// TIA Portal V20 export
TYPE "WT2_Vd_Status_1_UDT"
   STRUCT
      iHandshake : Int;
      Fehler : Struct
         bE0000_KonfigFehler : Bool;
         bE0001_VerbundMasterAusg : Bool;
         bE0002_NotstoppPHDFehler : Bool;
         bE0003_ExternFehler : Bool;
         bE0004_TDruckFehler : Bool;
         bE0005_PDruckFehler : Bool;
         bE0006_PSaugFehler : Bool;
         bE0007_TMotorFehler : Bool;
         bE0008_TSHMinSaugFehler : Bool;
         bE0009_TSHMinDruckFehler : Bool;
         bE0010_LuefterFehler : Bool;
         bE0011_Reserviert : Bool;
         bE0012_PhasenFehler : Bool;
         bE0013_MotorFehler : Bool;
         bE0014_LSAusloesung : Bool;
         bE0015_POeldiffStillstand : Bool;
         bE0016_POeldiffBetrieb : Bool;
         bE0017_TOelMaxFehler : Bool;
         bE0018_OElniveauOA : Bool;
         bE0019_OElniveauVd : Bool;
         bE0020_OElStroemung : Bool;
         bE0021_POelfilterBetrieb : Bool;
         bE0022_TLagerDEFehler : Bool;
         bE0023_TLager_NDEFehler : Bool;
         bE0024_Reserviert : Bool;
         bE0025_Reserviert : Bool;
         bE0026_Reserviert : Bool;
         bE0027_PSaugOverrange : Bool;
         bE0028_PPsZuTief : Bool;
         bE0029_Oelpumpe : Bool;
         bE0030_Leistungsschieber : Bool;
         bE0031_PoPsZuTief : Bool;
         bE0032_StartdruckZuHoch : Bool;
         bE0033_POelfilterStillstand : Bool;
         bE0034_PoPMinFehler : Bool;
         bE0035_Startoeldruck : Bool;
         bE0036_TDruckGradient : Bool;
         bE0037_OelflussVerdichter : Bool;
         bE0038_KeineGasfoerderung : Bool;
         bE0039_PZwDruck : Bool;
         bE0040_TZwDruck : Bool;
         bE0041_TSHMinZwDruck : Bool;
         bE0042_POeldiffMax : Bool;
         bE0043_PPsMax : Bool;
         bE0044_OelkhlungTop : Bool;
         bE0045_PPzZuTeif : Bool;
         bE0046_PPzMax : Bool;
         bE0047_PPsZuTief : Bool;
         bE0048_FluessigSchlag : Bool;
         bE0049_Reserviert : Bool;
         bE0050_Reserviert : Bool;
         bE0051_Reserviert : Bool;
         bE0052_Reserviert : Bool;
         bE0053_Reserviert : Bool;
         bE0054_Reserviert : Bool;
         bE0055_Reserviert : Bool;
         bE0056_Reserviert : Bool;
         bE0057_Reserviert : Bool;
         bE0058_Reserviert : Bool;
         bE0059_Reserviert : Bool;
         bE0060_Reserviert : Bool;
         bE0061_Reserviert : Bool;
         bE0062_Reserviert : Bool;
         bE0063_KaeltekreisMasterAusgefa : Bool;
         bE0064_Reserviert : Bool;
         bE0065_KaelteKreisInvUngueltig : Bool;
         bE0066_OelkreisMasterAusgefa : Bool;
         bE0067_Reserviert : Bool;
         bE0068_OelKreisInvUngueltig : Bool;
         bE0069_SchmierdruckMin : Bool;
         bE0070_PPoMax : Bool;
         bE0071_Haupt_OeldruckMin : Bool;
         bE0072_Reserviert : Bool;
         bE0073_Reserviert : Bool;
         bE0074_Reserviert : Bool;
         bE0075_TZylinderkopfFehler : Bool;
         bE0076_VerdampferpumpeFehlerBet : Bool;
         bE0077_VerdampferpumpeFehlerSti : Bool;
         bE0078_NivHDAbschHochFehler : Bool;
         bE0079_NivEconomiserHochFehler : Bool;
         bE0080_Reserviert : Bool;
         bE0081_KonfFehlerKkStart_Stopp : Bool;
         bE0082_HDVerdAusgefallen : Bool;
         bE0083_NDVerdAusgefallen : Bool;
         bE0084_KeinStartbefehlKonf : Bool;
         bE0085_PzPsMax : Bool;
         bE0086_Reserviert : Bool;
         bE0087_VibraSwitchAusg : Bool;
         bE0088_TOelabschMax : Bool;
         bE0089_TOelMin : Bool;
         bE0090_Reserviert : Bool;
         bE0091_NDAbschNivHoch : Bool;
         bE0092_Sekundaerschieber : Bool;
         bE0093_Reserviert : Bool;
         bE0094_KonfigFehlerAbsKuehls : Bool;
         bE0095_Reserviert : Bool;
         bE0096_OelnivKGHhoch : Bool;
         bE0097_KonfigFehlerDIPrio : Bool;
         bE0098_Reserviert : Bool;
         bE0099_Reserviert : Bool;
         bE0100_Reserviert : Bool;
         bE0101_KonfigFehlerDrehzahl : Bool;
         bE0102_Reserviert : Bool;
         bE0103_PSaugHoch : Bool;
         bE0104_KonfigFehlerMotorleist : Bool;
         bE0105_FehlerEinsatzdiagr : Bool;
         bE0106_Reserviert : Bool;
         bE0107_Reserviert : Bool;
         bE0108_Reserviert : Bool;
         bE0109_MotorfehlerNotAusTest : Bool;
         bE0110_StirnspHauptrotorZGross : Bool;
         bE0111_StirnspHautprotorZKlein : Bool;
         bE0112_StirnspNebenrotorZGross : Bool;
         bE0113_StirnspNebenrotorZKlein : Bool;
         bE0114_THauptrotorDS : Bool;
         bE0115_THauptrotorSS : Bool;
         bE0116_TNebenrotorDS : Bool;
         bE0117_TNebenrotorSS : Bool;
         bE0118_FlSchlagFehlerSensor : Bool;
         bE0119_OelstoppventilFehler : Bool;
         bE0120_Reserviert : Bool;
         bE0121_Reserviert : Bool;
         bE0122_Reserviert : Bool;
         bE0123_Reserviert : Bool;
         bE0124_Reserviert : Bool;
         bE0125_Reserviert : Bool;
         bE0126_Reserviert : Bool;
         bE0127_Reserviert : Bool;
      END_STRUCT;
      Alarm : Struct
         bA1000_Reserviert : Bool;
         bA1001_VerbundMasterAusg : Bool;
         bA1002_Reserviert : Bool;
         bA1003_Reserviert : Bool;
         bA1004_TDruck : Bool;
         bA1005_PDruck : Bool;
         bA1006_Reserviert : Bool;
         bA1007_TMotor : Bool;
         bA1008_TSHMinSaug : Bool;
         bA1009_TSHMinDruck : Bool;
         bA1010_Reserviert : Bool;
         bA1011_Reserviert : Bool;
         bA1012_Reserviert : Bool;
         bA1013_Reserviert : Bool;
         bA1014_Reserviert : Bool;
         bA1015_Reserviert : Bool;
         bA1016_POeldiff_Betrieb : Bool;
         bA1017_TOelmax : Bool;
         bA1018_OelniveauOA : Bool;
         bA1019_Reserviert : Bool;
         bA1020_Reserviert : Bool;
         bA1021_POelfilterBetrieb : Bool;
         bA1022_TLagerDE : Bool;
         bA1023_TLagerNDE : Bool;
         bA1024_OelniveauOA_hoch : Bool;
         bA1025_Reserviert : Bool;
         bA1026_Reserviert : Bool;
         bA1027_PSaugOverrange : Bool;
         bA1028_PPszutief : Bool;
         bA1029_Reserviert : Bool;
         bA1030_Reserviert : Bool;
         bA1031_Reserviert : Bool;
         bA1032_Reserviert : Bool;
         bA1033_Reserviert : Bool;
         bA1034_PoPMin : Bool;
         bA1035_Reserviert : Bool;
         bA1036_Reserviert : Bool;
         bA1037_Reserviert : Bool;
         bA1038_Reserviert : Bool;
         bA1039_PZwDruck : Bool;
         bA1040_TZwDruck : Bool;
         bA1041_TSHminZwDruck : Bool;
         bA1042_Reserviert : Bool;
         bA1043_PPsmax : Bool;
         bA1044_Reserviert : Bool;
         bA1045_PPzzutief : Bool;
         bA1046_PPzmax : Bool;
         bA1047_PPszutief2 : Bool;
         bA1048_FluessigSchlag : Bool;
         bA1049_NDPendel : Bool;
         bA1050_TOelMin : Bool;
         bA1051_Reserviert : Bool;
         bA1052_OelheizungOA : Bool;
         bA1053_TSaug : Bool;
         bA1054_PSauglimit : Bool;
         bA1055_PDrucklimit : Bool;
         bA1056_LastabwurfMotorstrom : Bool;
         bA1057_MinLeistungnErr : Bool;
         bA1058_MaxLeistungnErr : Bool;
         bA1059_BalanceFNorm : Bool;
         bA1060_PrimaerschMaxNErr : Bool;
         bA1061_LastabwurfMotorleistung : Bool;
         bA1062_OelheizungKGH : Bool;
         bA1063_KaeltekreisMasterAusgef : Bool;
         bA1064_KaeltekreisSlaveAusgef : Bool;
         bA1065_Reserviert : Bool;
         bA1066_Reserviert : Bool;
         bA1067_OelkreisSlaveAusgef : Bool;
         bA1068_Reserviert : Bool;
         bA1069_SchmierdruckMin : Bool;
         bA1070_PPoMax : Bool;
         bA1071_HauptOeldruckMin : Bool;
         bA1072_Oelnachspeisung : Bool;
         bA1073_KdMasterAusgef : Bool;
         bA1074_VrMasterAusgef : Bool;
         bA1075_TZylinderkopf : Bool;
         bA1076_Reserviert : Bool;
         bA1077_Reserviert : Bool;
         bA1078_Reserviert : Bool;
         bA1079_Reserviert : Bool;
         bA1080_KdMasterAusef : Bool;
         bA1081_Reserviert : Bool;
         bA1082_Reserviert : Bool;
         bA1083_Reserviert : Bool;
         bA1084_Reserviert : Bool;
         bA1085_PzPsAlarm : Bool;
         bA1086_HauptMasterAusgef : Bool;
         bA1087_Reserviert : Bool;
         bA1088_TOelabschMaxAlarm : Bool;
         bA1089_TOelMinAlarm : Bool;
         bA1090_OelpumpePendelalarm : Bool;
         bA1091_Reserviert : Bool;
         bA1092_Reserviert : Bool;
         bA1093_TOelMinAlarmKGH : Bool;
         bA1094_Reserviert : Bool;
         bA1095_TZwDruckSaugHDAlarm : Bool;
         bA1096_OelniveauKGHHoch : Bool;
         bA1097_Reserviert : Bool;
         bA1098_MKaeltekrMasterAktiv : Bool;
         bA1099_MOelkreisMasterAktiv : Bool;
         "bA1100_Objekt-ID mehrfach vorhanden" : Bool;
         bA1101_Reserviert : Bool;
         bA1102_RekalibrierungMinNDurchg : Bool;
         bA1103_Reserviert : Bool;
         bA1104_Reserviert : Bool;
         bA1105_AlarmEinsatzdiagr : Bool;
         bA1106_AlarmEcoNivEndsch : Bool;
         bA1107_OelnachspDVrGesp : Bool;
         bA1108_OerektDVrGesp : Bool;
         bA1109_NotAusTestFehlgeschl : Bool;
         bA1110_StirnspHauptrotorZGross : Bool;
         bA1111_StirnspHauptrotorZKlein : Bool;
         bA1112_StirnspNebenrotorZGross : Bool;
         bA1113_StirnspNebenrotorZKlein : Bool;
         bA1114_THauptrotorDS : Bool;
         bA1115_THauptrotorSS : Bool;
         bA1116_TNebenrotorDS : Bool;
         bA1117_TNebenrotorSS : Bool;
         bA1118_FlSchlagAlarmSensor : Bool;
         bA1119_Reserviert : Bool;
         bA1120_PDruckMinAlarm : Bool;
         bA1121_Vorschm10Tagen : Bool;
         bA1122_Vorschm9Tagen : Bool;
         bA1123_Vorschm8Tagen : Bool;
         bA1124_Vorschm7Tagen : Bool;
         bA1125_Vorschm6Tagen : Bool;
         bA1126_Vorschm5Tagen : Bool;
         bA1127_Vorschm4Tagen : Bool;
      END_STRUCT;
      Zustand : Struct
         bFehlerzustandAktiv : Bool;
         bAlarmzustandAktiv : Bool;
         bSystemMeldungAktiv : Bool;
         bServiceMeldungAktiv : Bool;
         bStopManuell : Bool;
         bStopAuto : Bool;
         bStopExtern : Bool;
         bBetriebAuto : Bool;
         bBetriebManuell : Bool;
         bAnlaufAuto : Bool;
         bAnlaufManuell : Bool;
         bManuellStoppen : Bool;
         b354_Reserve : Bool;
         b355_Reserve : Bool;
         b356_Reserve : Bool;
         b357_Reserve : Bool;
         by36_Reserve : Byte;
         bAnlaufsperre : Bool;
         bVerdichterSaugtAb : Bool;
         bLastabwurfSaugseite : Bool;
         bLastabwurfDruckseite : Bool;
         bLastabwurfPPs : Bool;
         bElStromGrNormal : Bool;
         bElStromGrMaximum : Bool;
         bOelZuKalt : Bool;
         bNiveauOelabschZuTief : Bool;
         bExternsperreAktiv : Bool;
         bEnergiesperreAktiv : Bool;
         bFreigabeWeitVdFehlt : Bool;
         bExternLimitAktiv : Bool;
         bInternLimitAktiv : Bool;
         bVerdichterVollOel : Bool;
         bOelabscheiderProblem : Bool;
         bBegrenzungElStromAktiv : Bool;
         bSealLube : Bool;
         bKeineFrgZwischendruck : Bool;
         bElLeistungGrNormal : Bool;
         bElLeistungGrMaximum : Bool;
         bBegrElLeistungAkt : Bool;
         bStartbefehlManuell : Bool;
         bOelpumpeManuell : Bool;
         bOelrektifizierungMan : Bool;
         bOelkuehlerManuell : Bool;
         bInventarKaeltekreis : Bool;
         bInventarOelkreis : Bool;
         bMasterGesperrt : Bool;
         bKaeltekrStbyMstInit : Bool;
         bKaeltekrStbyMstPassiv : Bool;
         bKaeltekrStbyMstAktiv : Bool;
         bHaltManuell : Bool;
         bGespVomKd : Bool;
         bGespVomVr : Bool;
         bOelZuWarm : Bool;
         bNachkalMin : Bool;
         bPDruckZuHoch : Bool;
         bVdStartVerz : Bool;
         bSchieberZwangstr : Bool;
         bGespVonOelkreisMaster : Bool;
         b421_Reserve : Bool;
         b422_Reserve : Bool;
         b423_Reserve : Bool;
         b424_Reserve : Bool;
         b425_Reserve : Bool;
         b426_Reserve : Bool;
         b427_Reserve : Bool;
         by43_Reserve : Byte;
         by44_Reserve : Byte;
         by45_Reserve : Byte;
      END_STRUCT;
      DigIn : Struct
         bNotstopp : Bool;
         bFehlerExtern : Bool;
         bPhasenuberwachung : Bool;
         bNiveauOelabscheiderTief : Bool;
         bNiveauOelabscheiderHoch : Bool;
         bNiveauKurbelgehaeuseTief : Bool;
         bNiveauOelabscheiderRueckf : Bool;
         bStartbefehl : Bool;
         bRmVerdichtermotor : Bool;
         bRmElOelpumpe : Bool;
         bExternLeistungslimit : Bool;
         bStartprioritaet : Bool;
         bRmChillerpumpe : Bool;
         bSpitzenlastsperre : Bool;
         bMotorbegrenzung : Bool;
         bPDruckseiteDigital : Bool;
         bPSaugseiteDigital : Bool;
         bPOelLubeDigital : Bool;
         bPOelfilterDigital : Bool;
         bTDruckseiteDigital : Bool;
         bTSaugseiteDigital : Bool;
         bTOelDigital : Bool;
         bTOelabscheiderDigital : Bool;
         bTMotorDigital : Bool;
         bNivKurbelGehaeuseHoch : Bool;
         bRueckmeldungLuefter : Bool;
         bRueckmeldungStoerung : Bool;
         bNivNDAbschHoch : Bool;
         bNivEconomiserHoch : Bool;
         bLastsperre : Bool;
         b496_Reserviert : Bool;
         bOelstrBitzer : Bool;
         bOelflussYork : Bool;
         bOelabschNivNormal : Bool;
         bAuxDigital1 : Bool;
         bAuxDigital2 : Bool;
         bVerdichterOelniveau : Bool;
         bVibraSwitch : Bool;
         bNDAbschNiveauHochMax : Bool;
         bStartzwangExtern : Bool;
         bOelnivKurbelGehaeuseNorm : Bool;
         bExternsperre : Bool;
         bDrehmomentbegrenzung : Bool;
         bNiveauEconomOpen : Bool;
         bNiveauEconomClose : Bool;
         bOelstoppventilBitzer : Bool;
         bFreigabePDruckLimit : Bool;
         bFreigabePSaugLimit : Bool;
         bFreigabeHaltebetrieb : Bool;
         b521_Reserve : Bool;
         b522_Reserve : Bool;
         b523_Reserve : Bool;
         b524_Reserve : Bool;
         b525_Reserve : Bool;
         b526_Reserve : Bool;
         b527_Reserve : Bool;
         by53_Reserve : Byte;
      END_STRUCT;
      DigOut : Struct
         bFehler : Bool;
         bAlarm : Bool;
         bLastschalterAusloesung : Bool;
         bBereit : Bool;
         bStart_Motor : Bool;
         bAnlaufentlastung : Bool;
         bTeilwicklung2 : Bool;
         bMagnetventilFluessig : Bool;
         bOelheizungOelabscheider : Bool;
         bOelheizungKurbelgehaeuse : Bool;
         bStartOelpumpe : Bool;
         bOelventil : Bool;
         bOelrektifizierungA : Bool;
         bOelrektifizierungB : Bool;
         bOelrueckfuehrung : Bool;
         bOelnachspeisung : Bool;
         bOelkuehlung : Bool;
         bPowerkit : Bool;
         bEconomiser : Bool;
         bLeistungGrGrenzwert : Bool;
         bZwischendruckkuehlung : Bool;
         bVerdapferpumpe : Bool;
         bStartanzeige : Bool;
         bGrundlastzylinder : Bool;
         bViMax : Bool;
         bViMin : Bool;
         bVi22 : Bool;
         bVi2235 : Bool;
         bUeberhitzungsventil : Bool;
         bStillstandentlastung : Bool;
         bOeltransfer : Bool;
         bFastPullDownMV : Bool;
         bNiveaureglerEconom : Bool;
         bOelrektEinzeln : Bool;
         bSaugleitungsheizung : Bool;
         bLeistungsschPulsBitzer : Bool;
         bAnzSchmierungNStillstand : Bool;
         bTOPHeizung : Bool;
         bTOPMVKuehlen : Bool;
         b587_Reserve : Bool;
         by59_Reserve : Byte;
         by60_Reserve : Byte;
         by61_Reserve : Byte;
      END_STRUCT;
      rPDruckBar : Real;
      rPDruckGrad : Real;
      rPSaugBar : Real;
      rPSaugGrad : Real;
      rIstleistProz : Real;
      rIstleistVol : Real;
      rSollleistProz : Real;
      rSollleistVol : Real;
      rIstVi : Real;
      rSollVi : Real;
      rPZwStufeBar : Real;
      rPZwStufeGrad : Real;
      rPEcoBar : Real;
      rPEcoGrad : Real;
      rPOelLube : Real;
      rPOelDiff : Real;
      rPOelfilter : Real;
      rPOelpumpe : Real;
      rPKGH : Real;
      rTDruck : Real;
      rTSaug : Real;
      rTZwStufe : Real;
      rTOel : Real;
      rTOelabscheider : Real;
      rTSHDruck : Real;
      rTSHSaug : Real;
      rTSHZwStufe : Real;
      rMotorstromA : Real;
      rMotorstromProz : Real;
      rMotorleistkW : Real;
      rMotorleistProz : Real;
      rMotorPTC : Real;
      diEinschaltMotor : DInt;
      diBetriebsstunden : DInt;
      iAktVdStufe : Int;
      rOelkRegIst : Real;
      rOelkRegSoll : Real;
      rOelkRegOut : Real;
      rMotordrehzahl : Real;
      diEnergiezaehlerTot : DInt;
      rOaNiveau : Real;
      rAuxAnalog1 : Real;
      rMinLeistung : Real;
      rMaxLeistung : Real;
      rPOelfilterEinAus : Real;
      rTOelkuehlerEin : Real;
      rTOelkuehlerAus : Real;
      rPosPriSchieber : Real;
      rPosSekSchieber : Real;
      rTSaugleitung : Real;
      rReserveReal : Array[0..14] of Real;
   END_STRUCT;
END_TYPE
